// TIA Portal V15.1 export
// export: Created 2026-11-02T18:55:11.1946213Z, ExportSetting WithDefaults, DisplayName Totally Integrated Automation Portal, DisplayVersion V15.1, DisplayName TIA Portal Openness, DisplayVersion V15.1, DisplayName STEP 7 Professional, DisplayVersion V15.1, DisplayName WinCC Professional, DisplayVersion V15.1
DATA_BLOCK "BR01_DB"   // DB3
{ S7_Optimized_Access := 'TRUE' }
VERSION : 0.1
// stored: AutoNumber false, InstanceOfName Burner, InstanceOfType FB
"Burner"
   // VAR_INPUT
   //    Auto : Bool;
   //    StartPB : Bool;
   //    StopOK : Bool;
   //    LevelOK : Bool;
   //    RunFb : Bool;
   //    Lockout : Bool;
   //    Fuel : Bool;
   //    TeA : Int;
   //    TeB : Int;
   //    Use24h : Bool;
   //    EStopOK : Bool;
   //    ResetPulse : Bool;
   //    FirstScan : Bool;
   //    SP : Int;
   //    HYST : Int;
   //    STG : Int;
   //    TStart : Time;
   // END_VAR
   // VAR_OUTPUT
   //    HeatReq : Bool;
   //    Stage2 : Bool;
   //    State : Int;
   //    Enabled : Bool;
   //    Tmax : Int;
   //    F_EStop : Bool;
   //    F_TC : Bool;
   //    F_Lockout : Bool;
   //    F_NoStart : Bool;
   //    F_RunLost : Bool;
   //    F_RunWrong : Bool;
   //    ParPending : Bool;
   // END_VAR
   // VAR
   //    StartEdge : Bool;
   //    StartMem : Bool;
   //    AutoChg : Bool;
   //    AutoMem : Bool;
   //    FuelChg : Bool;
   //    FuelMem : Bool;
   //    TcOkA : Bool;
   //    TcOkB : Bool;
   //    TcOk : Bool;
   //    TcBad : Bool;
   //    Demand : Bool;
   //    HeatNeed : Bool;
   //    Ready : Bool;
   //    Active : Bool;
   //    Pause24 : Bool;
   //    RunWrong : Bool;
   //    NoStart : Bool;
   //    PwrUpDone : Bool;
   //    TcSlow : Bool;
   //    SP_Act : Int;
   //    HYST_Act : Int;
   //    STG_Act : Int;
   //    TStart_Act : Time;
   //    TOn : Int;
   //    TStg : Int;
   //    TStgOff : Int;
   //    T_PwrUp : TON_TIME;
   //    T_TcBad : TON_TIME;
   //    T_24h : TON_TIME;
   //    T_Pause : TON_TIME;
   //    T_RunOff : TON_TIME;
   //    T_Start : TON_TIME;
   // END_VAR
BEGIN
END_DATA_BLOCK
